GLOBALCONSTANTS DialogIDs (* Objekt-IDs der Dialog-Vorlage *)
  (* Standard: 61499-2; Description: Copyright (c) 2026 Meisterschulen am Ostbahnhof This program and the accompanying materials are made available under the terms of the Eclipse Public License 2.0 which is available at https://www.eclipse.org/legal/epl-2.0/ SPDX-License-Identifier: EPL-2.0 *)
  (* Version 1.0, 2026-11-17, Franz Höpfinger, Meisterschulen am Ostbahnhof, initial API and implementation and/or initial documentation *)
  PACKAGE isobus::UT::dialog;
  VAR_GLOBAL CONSTANT
    Container_Dialog : UINT := UINT#3400; (* Vorlage Workspace_Dialog *)
    Container_Dlg_Box : UINT := UINT#3401; (* Vorlage Workspace_Dialog *)
    Rectangle_Dlg_Cover : UINT := UINT#14400; (* Vorlage Workspace_Dialog *)
    FillAttributes_Dlg_Title : UINT := UINT#25402; (* Vorlage Workspace_Dialog *)
    ObjectPointer_Dlg_Cover : UINT := UINT#27900; (* Vorlage Workspace_Dialog *)
    ObjectPointer_Dlg_Icon : UINT := UINT#27901; (* Vorlage Workspace_Dialog *)
    ObjectPointer_Dlg_Title : UINT := UINT#27902; (* Vorlage Workspace_Dialog *)
    ObjectPointer_Dlg_Text : UINT := UINT#27903; (* Vorlage Workspace_Dialog *)
    ObjectPointer_Dlg_Buttons : UINT := UINT#27904; (* Vorlage Workspace_Dialog *)
    Container_Dlg_Icon_Info : UINT := UINT#3402; (* Vorlage Workspace_Dialog *)
    Container_Dlg_Icon_Question : UINT := UINT#3403; (* Vorlage Workspace_Dialog *)
    Container_Dlg_Icon_Warning : UINT := UINT#3404; (* Vorlage Workspace_Dialog *)
    Container_Dlg_Icon_Error : UINT := UINT#3405; (* Vorlage Workspace_Dialog *)
    OutputString_Dlg_Title_Info : UINT := UINT#11410; (* Vorlage Workspace_Dialog *)
    OutputString_Dlg_Title_Question : UINT := UINT#11411; (* Vorlage Workspace_Dialog *)
    OutputString_Dlg_Title_Warning : UINT := UINT#11412; (* Vorlage Workspace_Dialog *)
    OutputString_Dlg_Title_Error : UINT := UINT#11413; (* Vorlage Workspace_Dialog *)
    Container_Dlg_Buttons_OK : UINT := UINT#3410; (* Vorlage Workspace_Dialog *)
    Container_Dlg_Buttons_OKCancel : UINT := UINT#3411; (* Vorlage Workspace_Dialog *)
    Container_Dlg_Buttons_AbortRetryIgnore : UINT := UINT#3412; (* Vorlage Workspace_Dialog *)
    Container_Dlg_Buttons_YesNoCancel : UINT := UINT#3413; (* Vorlage Workspace_Dialog *)
    Container_Dlg_Buttons_YesNo : UINT := UINT#3414; (* Vorlage Workspace_Dialog *)
    Container_Dlg_Buttons_RetryCancel : UINT := UINT#3415; (* Vorlage Workspace_Dialog *)
    Button_Dlg_OK : UINT := UINT#6900; (* Vorlage Workspace_Dialog *)
    Button_Dlg_Cancel : UINT := UINT#6901; (* Vorlage Workspace_Dialog *)
    Button_Dlg_Abort : UINT := UINT#6902; (* Vorlage Workspace_Dialog *)
    Button_Dlg_Retry : UINT := UINT#6903; (* Vorlage Workspace_Dialog *)
    Button_Dlg_Ignore : UINT := UINT#6904; (* Vorlage Workspace_Dialog *)
    Button_Dlg_Yes : UINT := UINT#6905; (* Vorlage Workspace_Dialog *)
    Button_Dlg_No : UINT := UINT#6906; (* Vorlage Workspace_Dialog *)
  END_VAR
END_GLOBALCONSTANTS
